// TIA Portal V19 export
TYPE "Pan_From_SM"
   STRUCT
      Supersaturation { ExternalWritable := 'False'} : Real;
      Crystal_Size { ExternalWritable := 'False'} : Real;
      Crystal_Content { ExternalWritable := 'False'} : Real;
      Mother_Liquor_Purity { ExternalWritable := 'False'} : Real;
      Concentration { ExternalWritable := 'False'} : Real;
      Temperature { ExternalWritable := 'False'} : Real;
      Refractometer_QF { ExternalWritable := 'False'} : Real;
      Massecuite_Solids_Content { ExternalWritable := 'False'} : Real;
      Density { ExternalWritable := 'False'} : Real;
      Steam_Valve_Control { ExternalWritable := 'False'} : Real;
      Vacuum_Valve_Control { ExternalWritable := 'False'} : Real;
      Syrup_Feed_Valve_Control { ExternalWritable := 'False'} : Real;
      real_reserve_1 : Real;
      real_reserve_2 : Real;
      real_reserve_3 : Real;
      real_reserve_4 : Real;
      real_reserve_5 : Real;
      Strike_Active { ExternalWritable := 'False'} : Bool;
      Seeded { ExternalWritable := 'False'} : Bool;
      Seeding_Valve_Control { ExternalWritable := 'False'} : Bool;
      Seeding_Warning { ExternalWritable := 'False'} : Bool;
      reserved_bit_48_4 { ExternalWritable := 'False'} : Bool;
      reserved_bit_48_5 { ExternalWritable := 'False'} : Bool;
      reserved_bit_48_6 { ExternalWritable := 'False'} : Bool;
      reserved_bit_48_7 { ExternalWritable := 'False'} : Bool;
   END_STRUCT;
END_TYPE
